TEXTLIST TextList_Piston_Recipe_State_CloseOpen
  0 = ' '
  1 = 'Close'
  2 = 'Open'
   = ''
END_TEXTLIST

(* stored: Version 1.1.0.1, ProductVersion 3.1.4024.12
   TextList TextList_Piston_Recipe_State_CloseOpen: Id {b3319678-2b43-4499-b67a-6ea6e5330180} *)
